(* IEC 61131-3 sources: Gen-AI/final/Gen-AI_v1.0_submission/A2_框架源码/agent/logs/full34_fixture/E3_S02_1_42/tools/candidate_1/fixture_compile, 1 file *)

(* ---- source.st ---- *)
FUNCTION_BLOCK FB_S02
VAR_INPUT
    FwdBtn : BOOL;
    RevBtn : BOOL;
    MaintKey : BOOL;
    EStop_NC : BOOL;
END_VAR
VAR_OUTPUT
    MotorFwd : BOOL;
    MotorRev : BOOL;
    RunLamp : BOOL;
    Status : WORD;
END_VAR
(* Add a VAR block for internal state/timers before the implementation, if needed. *)
(* SKELETON ONLY: replace this RETURN with scan logic and required initial state. *)
RETURN;
END_FUNCTION_BLOCK

(* FIXTURE_COMPILE_FAIL *)
